Fanuc KAREL source: KT00993.KL

PROGRAM KT00993
%NOLOCKGROUP
VAR
  P1: XYZWPREXT
  P2: XYZWPREXT
  X: REAL
  Y: REAL
  Z: REAL
  W: REAL
  P: REAL
  R: REAL
  CFG: CONFIG
BEGIN
  P1.X = 1.0
  P2.Y = 2.0
  P1.X = 1.0
  P2.Y = 2.0
  UNPOS(P1, X, Y, Z, W, P, R, CFG)
END KT00993
